# EPICS substitutions: db/Beckhoff_7XXX/ecmcEP7211-0034_OPT_encoder.substitutions
file "ecmcEL72XX_ENC.template"
{
  pattern {CH_ID}
          {01   }
}
